// ============================================================================
// DB_1006_ManualTeach_DJ005.scl - FB_1006_ManualTeach_BufferFraming 的背景数据块 (V15.1.0, 2026-11-15)
// ============================================================================
// 功能说明: 手动 / 示教。
//   背景 DB 不写变量, 变量来自 FB; 由 OB1 调用 "DB_1006_ManualTeach_DJ005"(...) 时使用。
//   TIA 全局 DB 里不能放 FB 实例, 故每个功能块一个背景 DB (LSP-905 §4.11)。
// ============================================================================

DATA_BLOCK "DB_1006_ManualTeach_DJ005"
"FB_1006_ManualTeach_BufferFraming"
BEGIN
END_DATA_BLOCK
